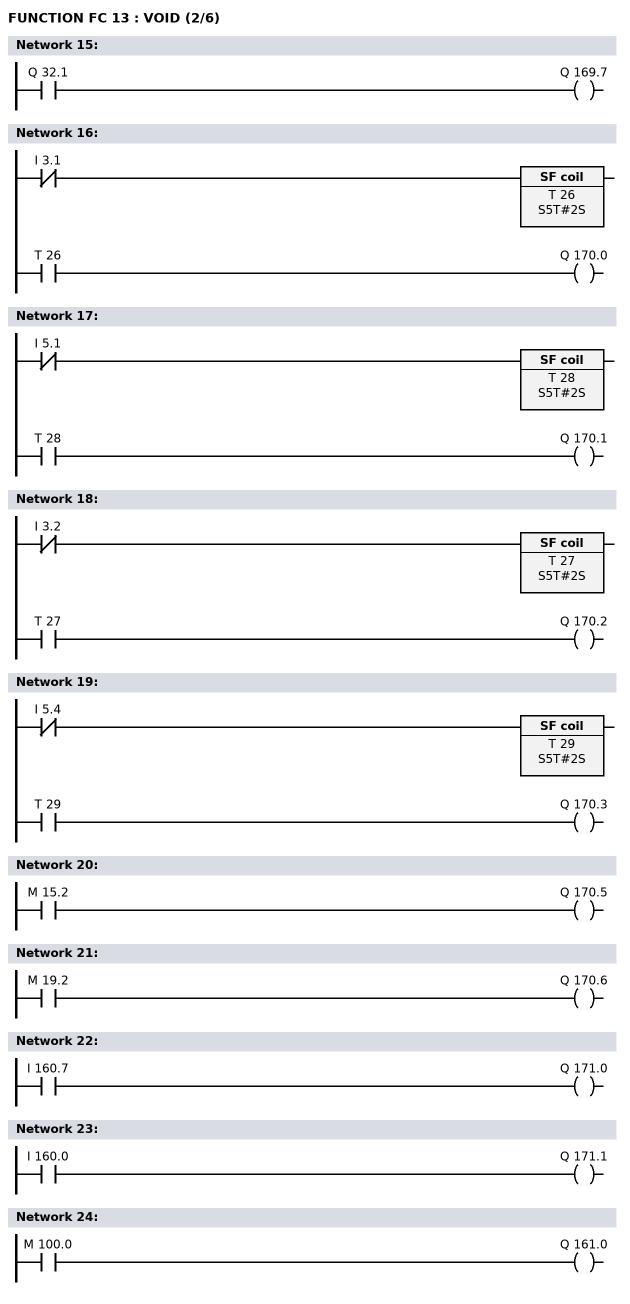

      A     Q     32.1;
      =     Q    169.7;
NETWORK
TITLE =

      AN    I      3.1;
      L     S5T#2S;
      SF    T     26;
      NOP   0;
      NOP   0;
      NOP   0;
      A     T     26;
      =     Q    170.0;
NETWORK
TITLE =

      AN    I      5.1;
      L     S5T#2S;
      SF    T     28;
      NOP   0;
      NOP   0;
      NOP   0;
      A     T     28;
      =     Q    170.1;
NETWORK
TITLE =

      AN    I      3.2;
      L     S5T#2S;
      SF    T     27;
      NOP   0;
      NOP   0;
      NOP   0;
      A     T     27;
      =     Q    170.2;
NETWORK
TITLE =

      AN    I      5.4;
      L     S5T#2S;
      SF    T     29;
      NOP   0;
      NOP   0;
      NOP   0;
      A     T     29;
      =     Q    170.3;
NETWORK
TITLE =

      A     M     15.2;
      =     Q    170.5;
NETWORK
TITLE =

      A     M     19.2;
      =     Q    170.6;
NETWORK
TITLE =

      A     I    160.7;
      =     Q    171.0;
NETWORK
TITLE =

      A     I    160.0;
      =     Q    171.1;
NETWORK
TITLE =

      A     M    100.0;
      =     Q    161.0;
NETWORK
TITLE =
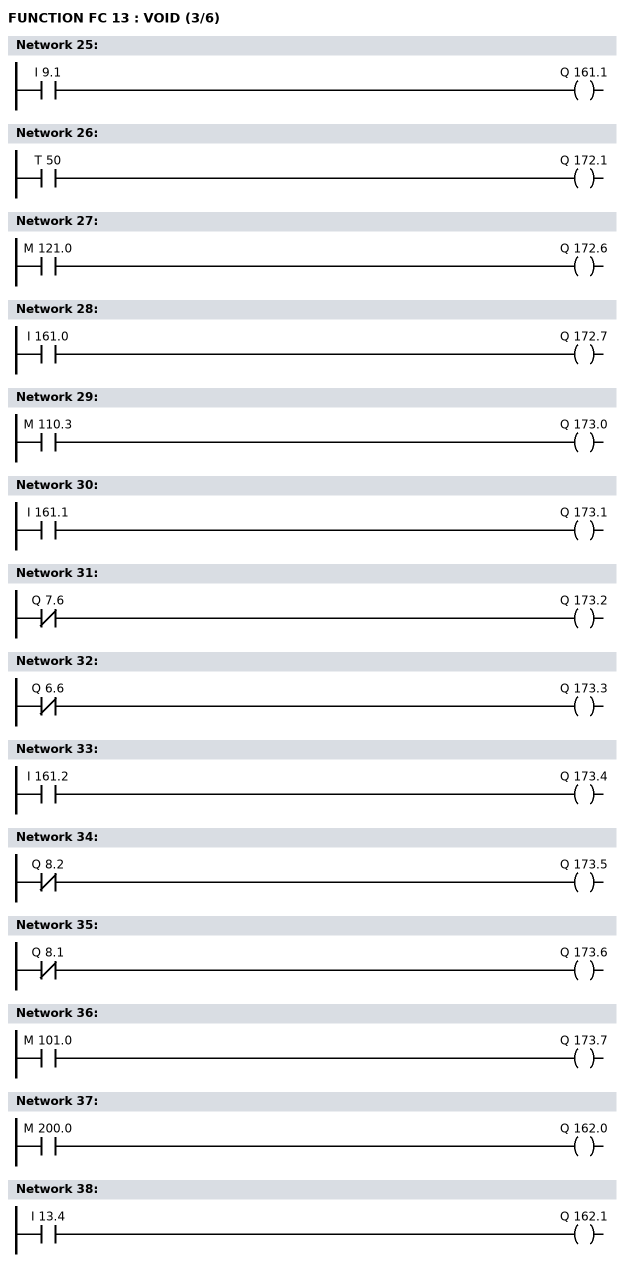

      A     I      9.1;
      =     Q    161.1;
NETWORK
TITLE =

      A     T     50;
      =     Q    172.1;
NETWORK
TITLE =

      A     M    121.0;
      =     Q    172.6;
NETWORK
TITLE =

      A     I    161.0;
      =     Q    172.7;
NETWORK
TITLE =

      A     M    110.3;
      =     Q    173.0;
NETWORK
TITLE =

      A     I    161.1;
      =     Q    173.1;
NETWORK
TITLE =

      AN    Q      7.6;
      =     Q    173.2;
NETWORK
TITLE =

      AN    Q      6.6;
      =     Q    173.3;
NETWORK
TITLE =

      A     I    161.2;
      =     Q    173.4;
NETWORK
TITLE =

      AN    Q      8.2;
      =     Q    173.5;
NETWORK
TITLE =

      AN    Q      8.1;
      =     Q    173.6;
NETWORK
TITLE =

      A     M    101.0;
      =     Q    173.7;
NETWORK
TITLE =

      A     M    200.0;
      =     Q    162.0;
NETWORK
TITLE =

      A     I     13.4;
      =     Q    162.1;
NETWORK
TITLE =
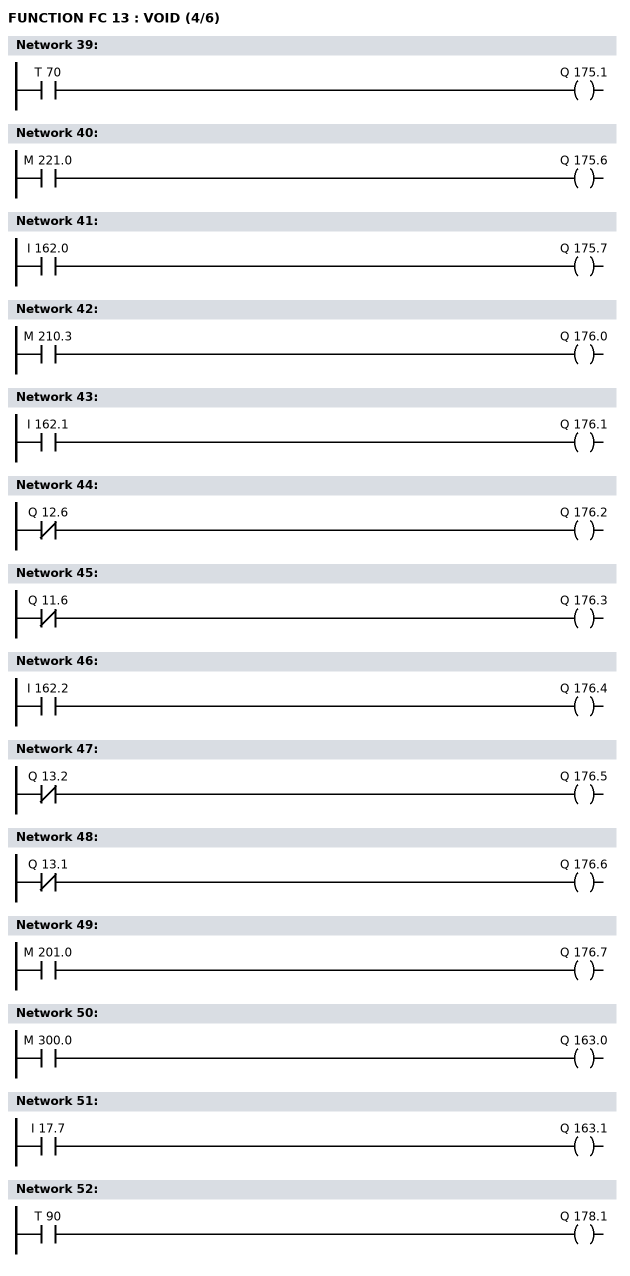

      A     T     70;
      =     Q    175.1;
NETWORK
TITLE =

      A     M    221.0;
      =     Q    175.6;
NETWORK
TITLE =

      A     I    162.0;
      =     Q    175.7;
NETWORK
TITLE =

      A     M    210.3;
      =     Q    176.0;
NETWORK
TITLE =

      A     I    162.1;
      =     Q    176.1;
NETWORK
TITLE =

      AN    Q     12.6;
      =     Q    176.2;
NETWORK
TITLE =

      AN    Q     11.6;
      =     Q    176.3;
NETWORK
TITLE =

      A     I    162.2;
      =     Q    176.4;
NETWORK
TITLE =

      AN    Q     13.2;
      =     Q    176.5;
NETWORK
TITLE =

      AN    Q     13.1;
      =     Q    176.6;
NETWORK
TITLE =

      A     M    201.0;
      =     Q    176.7;
NETWORK
TITLE =

      A     M    300.0;
      =     Q    163.0;
NETWORK
TITLE =

      A     I     17.7;
      =     Q    163.1;
NETWORK
TITLE =

      A     T     90;
      =     Q    178.1;
NETWORK
TITLE =
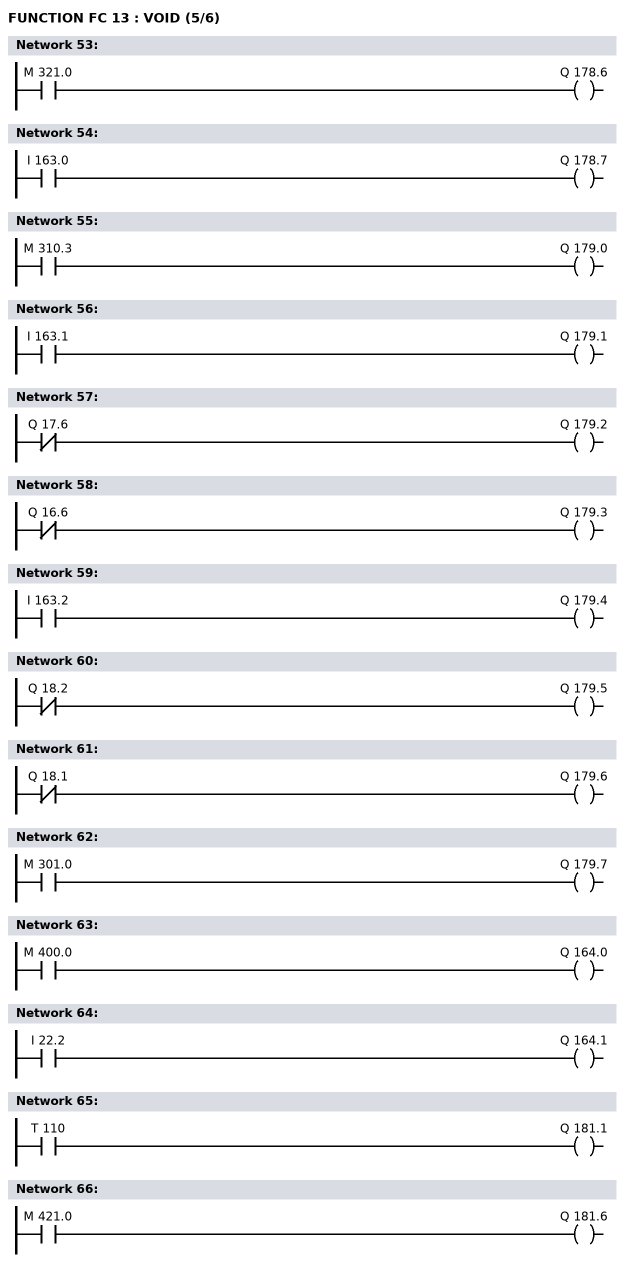

      A     M    321.0;
      =     Q    178.6;
NETWORK
TITLE =

      A     I    163.0;
      =     Q    178.7;
NETWORK
TITLE =

      A     M    310.3;
      =     Q    179.0;
NETWORK
TITLE =

      A     I    163.1;
      =     Q    179.1;
NETWORK
TITLE =

      AN    Q     17.6;
      =     Q    179.2;
NETWORK
TITLE =

      AN    Q     16.6;
      =     Q    179.3;
NETWORK
TITLE =

      A     I    163.2;
      =     Q    179.4;
NETWORK
TITLE =

      AN    Q     18.2;
      =     Q    179.5;
NETWORK
TITLE =

      AN    Q     18.1;
      =     Q    179.6;
NETWORK
TITLE =

      A     M    301.0;
      =     Q    179.7;
NETWORK
TITLE =

      A     M    400.0;
      =     Q    164.0;
NETWORK
TITLE =

      A     I     22.2;
      =     Q    164.1;
NETWORK
TITLE =

      A     T    110;
      =     Q    181.1;
NETWORK
TITLE =

      A     M    421.0;
      =     Q    181.6;
NETWORK
TITLE =
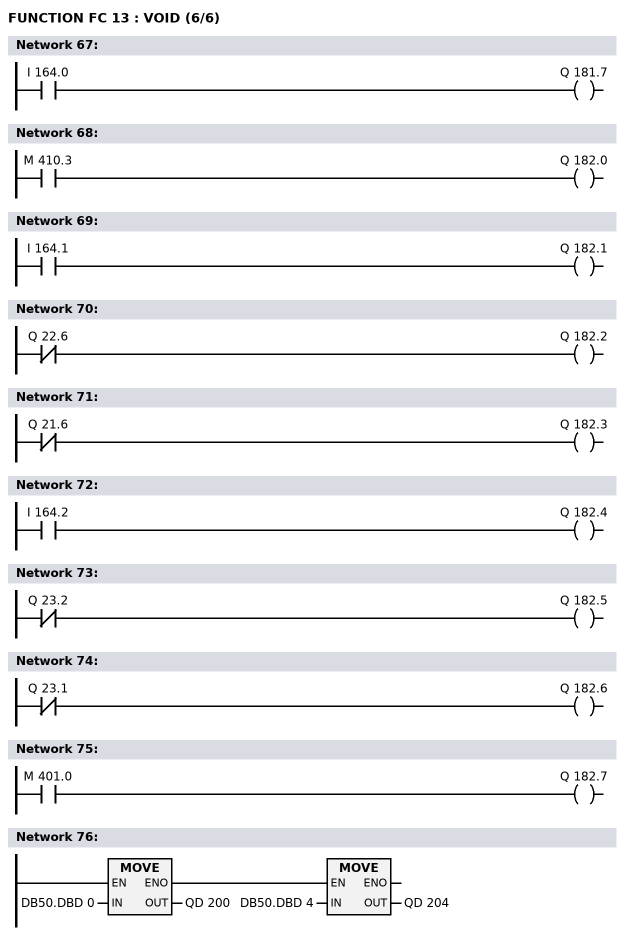

      A     I    164.0;
      =     Q    181.7;
NETWORK
TITLE =

      A     M    410.3;
      =     Q    182.0;
NETWORK
TITLE =

      A     I    164.1;
      =     Q    182.1;
NETWORK
TITLE =

      AN    Q     22.6;
      =     Q    182.2;
NETWORK
TITLE =

      AN    Q     21.6;
      =     Q    182.3;
NETWORK
TITLE =

      A     I    164.2;
      =     Q    182.4;
NETWORK
TITLE =

      AN    Q     23.2;
      =     Q    182.5;
NETWORK
TITLE =

      AN    Q     23.1;
      =     Q    182.6;
NETWORK
TITLE =

      A     M    401.0;
      =     Q    182.7;
NETWORK
TITLE =

      A(    ;
      L     DB50.DBD    0;
      T     QD   200;
      SET   ;
      SAVE  ;
      CLR   ;
      A     BR;
      )     ;
      JNB   M001;
      L     DB50.DBD    4;
      T     QD   204;
M001: NOP   0;
END_FUNCTION

FUNCTION FC 100 : VOID
VERSION : 0.1

BEGIN
NETWORK
TITLE =
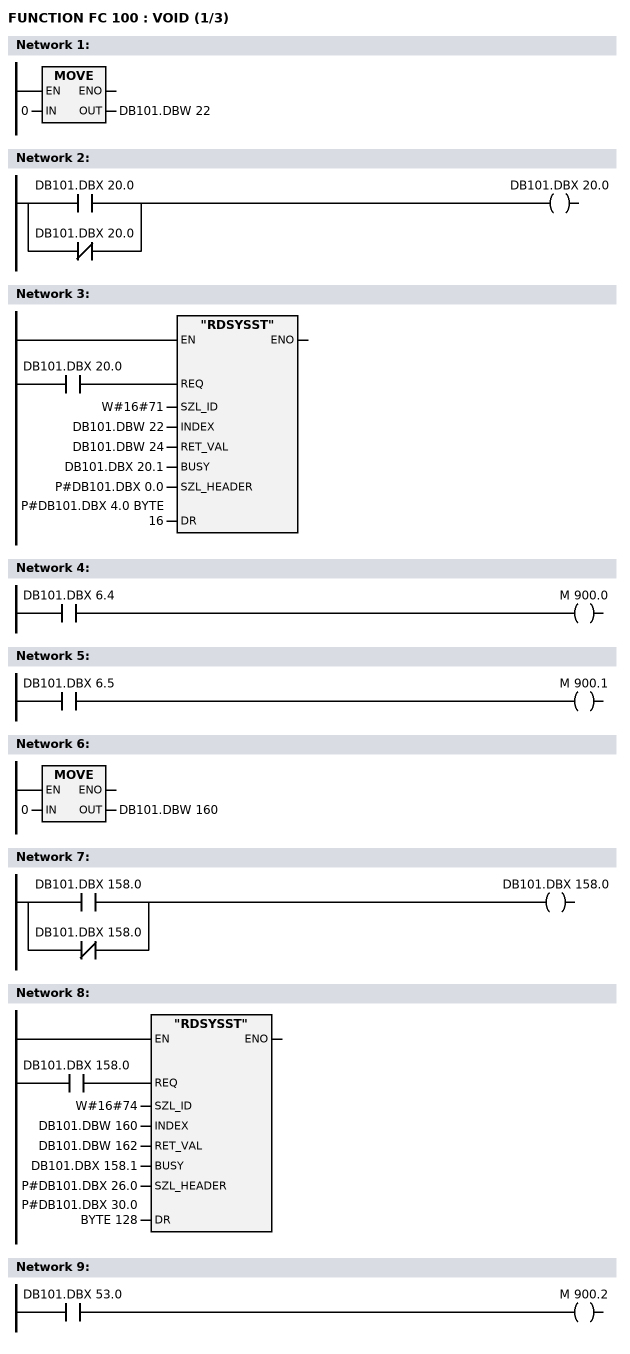

      L     0;
      T     DB101.DBW   22;
      NOP   0;
NETWORK
TITLE =

      O     DB101.DBX   20.0;
      ON    DB101.DBX   20.0;
      =     DB101.DBX   20.0;
NETWORK
TITLE =

      A     DB101.DBX   20.0;
      =     L      0.0;
      BLD   103;
      CALL "RDSYSST" (
           REQ                      := L      0.0,
           SZL_ID                   := W#16#71,
           INDEX                    := DB101.DBW   22,
           RET_VAL                  := DB101.DBW   24,
           BUSY                     := DB101.DBX   20.1,
           SZL_HEADER               := P#DB101.DBX 0.0,
           DR                       := P#DB101.DBX 4.0 BYTE 16);
      NOP   0;
NETWORK
TITLE =

      A     DB101.DBX    6.4;
      =     M    900.0;
NETWORK
TITLE =

      A     DB101.DBX    6.5;
      =     M    900.1;
NETWORK
TITLE =

      L     0;
      T     DB101.DBW  160;
      NOP   0;
NETWORK
TITLE =

      O     DB101.DBX  158.0;
      ON    DB101.DBX  158.0;
      =     DB101.DBX  158.0;
NETWORK
TITLE =

      A     DB101.DBX  158.0;
      =     L      0.0;
      BLD   103;
      CALL "RDSYSST" (
           REQ                      := L      0.0,
           SZL_ID                   := W#16#74,
           INDEX                    := DB101.DBW  160,
           RET_VAL                  := DB101.DBW  162,
           BUSY                     := DB101.DBX  158.1,
           SZL_HEADER               := P#DB101.DBX 26.0,
           DR                       := P#DB101.DBX 30.0 BYTE 128);
      NOP   0;
NETWORK
TITLE =

      A     DB101.DBX   53.0;
      =     M    900.2;
NETWORK
TITLE =
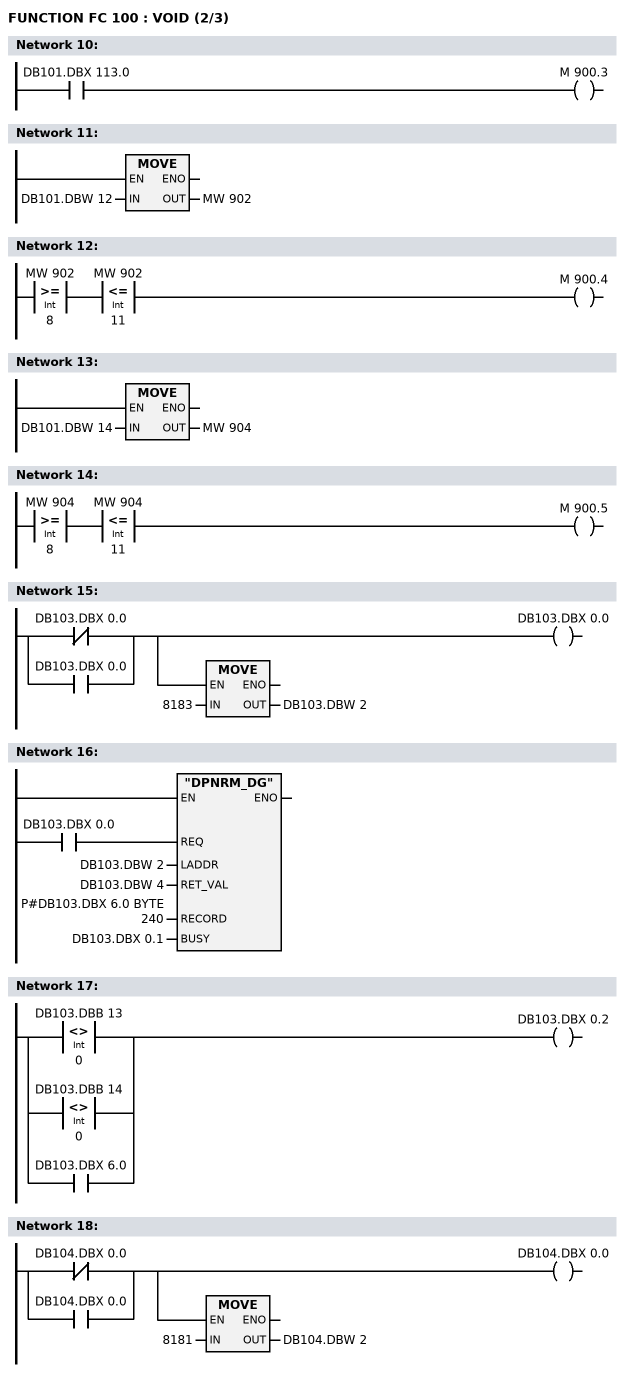

      A     DB101.DBX  113.0;
      =     M    900.3;
NETWORK
TITLE =

      L     DB101.DBW   12;
      T     MW   902;
      NOP   0;
NETWORK
TITLE =

      A(    ;
      L     MW   902;
      L     8;
      >=I   ;
      )     ;
      A(    ;
      L     MW   902;
      L     11;
      <=I   ;
      )     ;
      =     M    900.4;
NETWORK
TITLE =

      L     DB101.DBW   14;
      T     MW   904;
      NOP   0;
NETWORK
TITLE =

      A(    ;
      L     MW   904;
      L     8;
      >=I   ;
      )     ;
      A(    ;
      L     MW   904;
      L     11;
      <=I   ;
      )     ;
      =     M    900.5;
NETWORK
TITLE =

      ON    DB103.DBX    0.0;
      O     DB103.DBX    0.0;
      =     L      0.0;
      A     L      0.0;
      BLD   102;
      =     DB103.DBX    0.0;
      A     L      0.0;
      JNB   M001;
      L     8183;
      T     DB103.DBW    2;
M001: NOP   0;
NETWORK
TITLE =

      A     DB103.DBX    0.0;
      =     L      0.0;
      BLD   103;
      CALL "DPNRM_DG" (
           REQ                      := L      0.0,
           LADDR                    := DB103.DBW    2,
           RET_VAL                  := DB103.DBW    4,
           RECORD                   := P#DB103.DBX 6.0 BYTE 240,
           BUSY                     := DB103.DBX    0.1);
      NOP   0;
NETWORK
TITLE =

      O(    ;
      L     DB103.DBB   13;
      L     0;
      <>I   ;
      )     ;
      O(    ;
      L     DB103.DBB   14;
      L     0;
      <>I   ;
      )     ;
      O     DB103.DBX    6.0;
      =     DB103.DBX    0.2;
NETWORK
TITLE =

      ON    DB104.DBX    0.0;
      O     DB104.DBX    0.0;
      =     L      0.0;
      A     L      0.0;
      BLD   102;
      =     DB104.DBX    0.0;
      A     L      0.0;
      JNB   M002;
      L     8181;
      T     DB104.DBW    2;
M002: NOP   0;
NETWORK
TITLE =
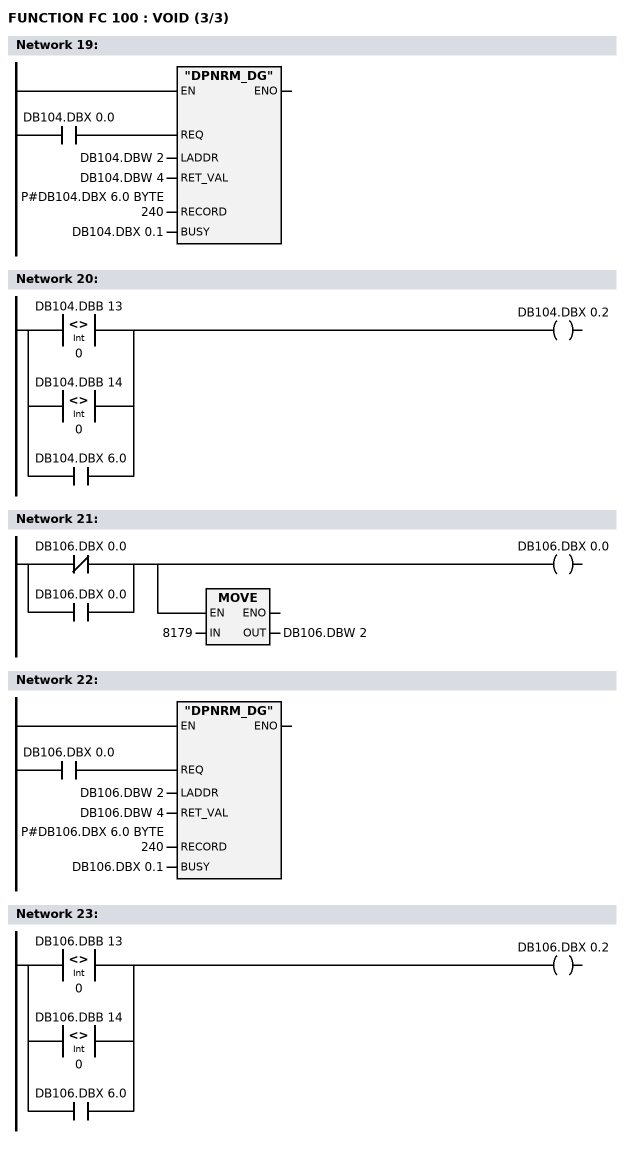

      A     DB104.DBX    0.0;
      =     L      0.0;
      BLD   103;
      CALL "DPNRM_DG" (
           REQ                      := L      0.0,
           LADDR                    := DB104.DBW    2,
           RET_VAL                  := DB104.DBW    4,
           RECORD                   := P#DB104.DBX 6.0 BYTE 240,
           BUSY                     := DB104.DBX    0.1);
      NOP   0;
NETWORK
TITLE =

      O(    ;
      L     DB104.DBB   13;
      L     0;
      <>I   ;
      )     ;
      O(    ;
      L     DB104.DBB   14;
      L     0;
      <>I   ;
      )     ;
      O     DB104.DBX    6.0;
      =     DB104.DBX    0.2;
NETWORK
TITLE =

      ON    DB106.DBX    0.0;
      O     DB106.DBX    0.0;
      =     L      0.0;
      A     L      0.0;
      BLD   102;
      =     DB106.DBX    0.0;
      A     L      0.0;
      JNB   M003;
      L     8179;
      T     DB106.DBW    2;
M003: NOP   0;
NETWORK
TITLE =

      A     DB106.DBX    0.0;
      =     L      0.0;
      BLD   103;
      CALL "DPNRM_DG" (
           REQ                      := L      0.0,
           LADDR                    := DB106.DBW    2,
           RET_VAL                  := DB106.DBW    4,
           RECORD                   := P#DB106.DBX 6.0 BYTE 240,
           BUSY                     := DB106.DBX    0.1);
      NOP   0;
NETWORK
TITLE =

      O(    ;
      L     DB106.DBB   13;
      L     0;
      <>I   ;
      )     ;
      O(    ;
      L     DB106.DBB   14;
      L     0;
      <>I   ;
      )     ;
      O     DB106.DBX    6.0;
      =     DB106.DBX    0.2;
END_FUNCTION

DATA_BLOCK DB 500
VERSION : 0.0

 FB 500
BEGIN
   IN0 := FALSE;
   IN1 := FALSE;
   IN2 := FALSE;
   OUT3 := FALSE;
   OUT4 := FALSE;
   STAT5 := FALSE;
   STAT6 := FALSE;
   STAT7 := FALSE;
   STAT8 := FALSE;
END_DATA_BLOCK

DATA_BLOCK DB 501
VERSION : 0.0

 FB 500
BEGIN
   IN0 := FALSE;
   IN1 := FALSE;
   IN2 := FALSE;
   OUT3 := FALSE;
   OUT4 := FALSE;
   STAT5 := FALSE;
   STAT6 := FALSE;
   STAT7 := FALSE;
   STAT8 := FALSE;
END_DATA_BLOCK

DATA_BLOCK DB 502
VERSION : 0.0

 FB 500
BEGIN
   IN0 := FALSE;
   IN1 := FALSE;
   IN2 := FALSE;
   OUT3 := FALSE;
   OUT4 := FALSE;
   STAT5 := FALSE;
   STAT6 := FALSE;
   STAT7 := FALSE;
   STAT8 := FALSE;
END_DATA_BLOCK

DATA_BLOCK DB 504
VERSION : 0.0

 FB 500
BEGIN
   IN0 := FALSE;
   IN1 := FALSE;
   IN2 := FALSE;
   OUT3 := FALSE;
   OUT4 := FALSE;
   STAT5 := FALSE;
   STAT6 := FALSE;
   STAT7 := FALSE;
   STAT8 := FALSE;
END_DATA_BLOCK

DATA_BLOCK DB 505
VERSION : 0.0

 FB 500
BEGIN
   IN0 := FALSE;
   IN1 := FALSE;
   IN2 := FALSE;
   OUT3 := FALSE;
   OUT4 := FALSE;
   STAT5 := FALSE;
   STAT6 := FALSE;
   STAT7 := FALSE;
   STAT8 := FALSE;
END_DATA_BLOCK

DATA_BLOCK DB 506
VERSION : 0.0

 FB 500
BEGIN
   IN0 := FALSE;
   IN1 := FALSE;
   IN2 := FALSE;
   OUT3 := FALSE;
   OUT4 := FALSE;
   STAT5 := FALSE;
   STAT6 := FALSE;
   STAT7 := FALSE;
   STAT8 := FALSE;
END_DATA_BLOCK

DATA_BLOCK DB 507
VERSION : 0.0

 FB 500
BEGIN
   IN0 := FALSE;
   IN1 := FALSE;
   IN2 := FALSE;
   OUT3 := FALSE;
   OUT4 := FALSE;
   STAT5 := FALSE;
   STAT6 := FALSE;
   STAT7 := FALSE;
   STAT8 := FALSE;
END_DATA_BLOCK

DATA_BLOCK DB 508
VERSION : 0.0

 FB 500
BEGIN
   IN0 := FALSE;
   IN1 := FALSE;
   IN2 := FALSE;
   OUT3 := FALSE;
   OUT4 := FALSE;
   STAT5 := FALSE;
   STAT6 := FALSE;
   STAT7 := FALSE;
   STAT8 := FALSE;
END_DATA_BLOCK

DATA_BLOCK DB 509
VERSION : 0.0

 FB 500
BEGIN
   IN0 := FALSE;
   IN1 := FALSE;
   IN2 := FALSE;
   OUT3 := FALSE;
   OUT4 := FALSE;
   STAT5 := FALSE;
   STAT6 := FALSE;
   STAT7 := FALSE;
   STAT8 := FALSE;
END_DATA_BLOCK

DATA_BLOCK DB 517
VERSION : 0.0

 FB 500
BEGIN
   IN0 := FALSE;
   IN1 := FALSE;
   IN2 := FALSE;
   OUT3 := FALSE;
   OUT4 := FALSE;
   STAT5 := FALSE;
   STAT6 := FALSE;
   STAT7 := FALSE;
   STAT8 := FALSE;
END_DATA_BLOCK

DATA_BLOCK DB 518
VERSION : 0.0

 FB 500
BEGIN
   IN0 := FALSE;
   IN1 := FALSE;
   IN2 := FALSE;
   OUT3 := FALSE;
   OUT4 := FALSE;
   STAT5 := FALSE;
   STAT6 := FALSE;
   STAT7 := FALSE;
   STAT8 := FALSE;
END_DATA_BLOCK

DATA_BLOCK DB 519
VERSION : 0.0

 FB 500
BEGIN
   IN0 := FALSE;
   IN1 := FALSE;
   IN2 := FALSE;
   OUT3 := FALSE;
   OUT4 := FALSE;
   STAT5 := FALSE;
   STAT6 := FALSE;
   STAT7 := FALSE;
   STAT8 := FALSE;
END_DATA_BLOCK

DATA_BLOCK DB 520
VERSION : 0.0

 FB 500
BEGIN
   IN0 := FALSE;
   IN1 := FALSE;
   IN2 := FALSE;
   OUT3 := FALSE;
   OUT4 := FALSE;
   STAT5 := FALSE;
   STAT6 := FALSE;
   STAT7 := FALSE;
   STAT8 := FALSE;
END_DATA_BLOCK

DATA_BLOCK DB 521
VERSION : 0.0

 FB 500
BEGIN
   IN0 := FALSE;
   IN1 := FALSE;
   IN2 := FALSE;
   OUT3 := FALSE;
   OUT4 := FALSE;
   STAT5 := FALSE;
   STAT6 := FALSE;
   STAT7 := FALSE;
   STAT8 := FALSE;
END_DATA_BLOCK

DATA_BLOCK DB 522
VERSION : 0.0

 FB 500
BEGIN
   IN0 := FALSE;
   IN1 := FALSE;
   IN2 := FALSE;
   OUT3 := FALSE;
   OUT4 := FALSE;
   STAT5 := FALSE;
   STAT6 := FALSE;
   STAT7 := FALSE;
   STAT8 := FALSE;
END_DATA_BLOCK

DATA_BLOCK DB 523
VERSION : 0.0

 FB 500
BEGIN
   IN0 := FALSE;
   IN1 := FALSE;
   IN2 := FALSE;
   OUT3 := FALSE;
   OUT4 := FALSE;
   STAT5 := FALSE;
   STAT6 := FALSE;
   STAT7 := FALSE;
   STAT8 := FALSE;
END_DATA_BLOCK

DATA_BLOCK DB 524
VERSION : 0.0

 FB 500
BEGIN
   IN0 := FALSE;
   IN1 := FALSE;
   IN2 := FALSE;
   OUT3 := FALSE;
   OUT4 := FALSE;
   STAT5 := FALSE;
   STAT6 := FALSE;
   STAT7 := FALSE;
   STAT8 := FALSE;
END_DATA_BLOCK

ORGANIZATION_BLOCK OB 1
VERSION : 0.1


VAR_TEMP
  TEMP0 : BYTE ;
  TEMP1 : BYTE ;
  TEMP2 : BYTE ;
  TEMP3 : BYTE ;
  TEMP4 : BYTE ;
  TEMP5 : BYTE ;
  TEMP6 : INT ;
  TEMP7 : INT ;
  TEMP8 : INT ;
  TEMP9 : DATE_AND_TIME ;
END_VAR
BEGIN
NETWORK
TITLE =
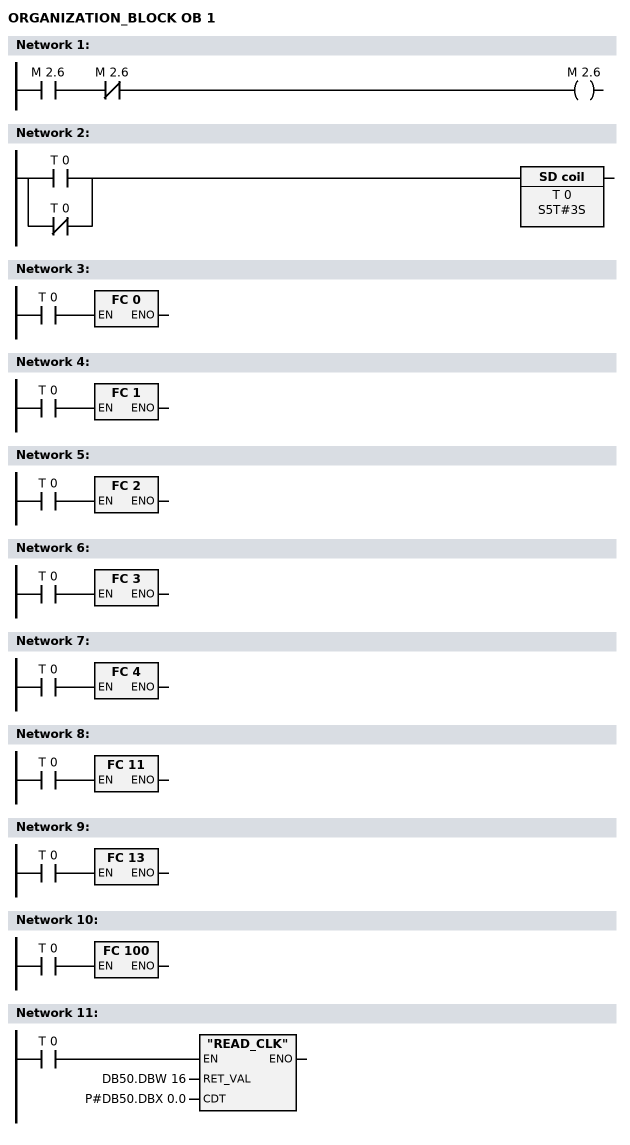

      A     M      2.6;
      AN    M      2.6;
      =     M      2.6;
NETWORK
TITLE =

      A(    ;
      O     T      0;
      ON    T      0;
      )     ;
      L     S5T#3S;
      SD    T      0;
      NOP   0;
      NOP   0;
      NOP   0;
      NOP   0;
NETWORK
TITLE =

      A     T      0;
      JNB   M001;
      CALL FC     0 ;
M001: NOP   0;
NETWORK
TITLE =

      A     T      0;
      JNB   M002;
      CALL FC     1 ;
M002: NOP   0;
NETWORK
TITLE =

      A     T      0;
      JNB   M003;
      CALL FC     2 ;
M003: NOP   0;
NETWORK
TITLE =

      A     T      0;
      JNB   M004;
      CALL FC     3 ;
M004: NOP   0;
NETWORK
TITLE =

      A     T      0;
      JNB   M005;
      CALL FC     4 ;
M005: NOP   0;
NETWORK
TITLE =

      A     T      0;
      JNB   M006;
      CALL FC    11 ;
M006: NOP   0;
NETWORK
TITLE =

      A     T      0;
      JNB   M007;
      CALL FC    13 ;
M007: NOP   0;
NETWORK
TITLE =

      A     T      0;
      JNB   M008;
      CALL FC   100 ;
M008: NOP   0;
NETWORK
TITLE =

      A     T      0;
      JNB   M009;
      CALL "READ_CLK" (
           RET_VAL                  := DB50.DBW   16,
           CDT                      := P#DB50.DBX 0.0);
M009: NOP   0;
END_ORGANIZATION_BLOCK

ORGANIZATION_BLOCK OB 35
VERSION : 0.1


VAR_TEMP
  TEMP0 : BYTE ;
  TEMP1 : BYTE ;
  TEMP2 : BYTE ;
  TEMP3 : BYTE ;
  TEMP4 : BYTE ;
  TEMP5 : BYTE ;
  TEMP6 : WORD ;
  TEMP7 : INT ;
  TEMP8 : INT ;
  TEMP9 : DATE_AND_TIME ;
END_VAR
BEGIN
END_ORGANIZATION_BLOCK

ORGANIZATION_BLOCK OB 70
VERSION : 0.1


VAR_TEMP
  TEMP0 : BYTE ;
  TEMP1 : BYTE ;
  TEMP2 : BYTE ;
  TEMP3 : BYTE ;
  TEMP4 : WORD ;
  TEMP5 : WORD ;
  TEMP6 : WORD ;
  TEMP7 : WORD ;
  TEMP8 : DATE_AND_TIME ;
END_VAR
BEGIN
NETWORK
TITLE =

      AN    M      3.7;
      =     M      3.7;
END_ORGANIZATION_BLOCK

ORGANIZATION_BLOCK OB 72
VERSION : 0.1


VAR_TEMP
  TEMP0 : BYTE ;
  TEMP1 : BYTE ;
  TEMP2 : BYTE ;
  TEMP3 : BYTE ;
  TEMP4 : WORD ;
  TEMP5 : WORD ;
  TEMP6 : WORD ;
  TEMP7 : WORD ;
  TEMP8 : DATE_AND_TIME ;
END_VAR
BEGIN
NETWORK
TITLE =

      A     M      3.7;
      =     M      3.7;
END_ORGANIZATION_BLOCK

ORGANIZATION_BLOCK OB 81
VERSION : 0.1


VAR_TEMP
  TEMP0 : BYTE ;
  TEMP1 : BYTE ;
  TEMP2 : BYTE ;
  TEMP3 : BYTE ;
  TEMP4 : BYTE ;
  TEMP5 : BYTE ;
  TEMP6 : WORD ;
  TEMP7 : BYTE ;
  TEMP8 : BYTE ;
  TEMP9 : BYTE ;
  TEMP10 : BYTE ;
  TEMP11 : DATE_AND_TIME ;
END_VAR
BEGIN
NETWORK
TITLE =

      AN    M      3.7;
      =     M      3.7;
END_ORGANIZATION_BLOCK

ORGANIZATION_BLOCK OB 82
VERSION : 0.1


VAR_TEMP
  TEMP0 : BYTE ;
  TEMP1 : BYTE ;
  TEMP2 : BYTE ;
  TEMP3 : BYTE ;
  TEMP4 : BYTE ;
  TEMP5 : BYTE ;
  TEMP6 : WORD ;
  TEMP7 : BOOL ;
  TEMP8 : BOOL ;
  TEMP9 : BOOL ;
  TEMP10 : BOOL ;
  TEMP11 : BOOL ;
  TEMP12 : BOOL ;
  TEMP13 : BOOL ;
  TEMP14 : BOOL ;
  TEMP15 : BYTE ;
  TEMP16 : BOOL ;
  TEMP17 : BOOL ;
  TEMP18 : BOOL ;
  TEMP19 : BOOL ;
  TEMP20 : BOOL ;
  TEMP21 : BOOL ;
  TEMP22 : BOOL ;
  TEMP23 : BOOL ;
  TEMP24 : BOOL ;
  TEMP25 : BOOL ;
  TEMP26 : BOOL ;
  TEMP27 : BOOL ;
  TEMP28 : BOOL ;
  TEMP29 : BOOL ;
  TEMP30 : BOOL ;
  TEMP31 : BOOL ;
  TEMP32 : DATE_AND_TIME ;
END_VAR
BEGIN
NETWORK
TITLE =

      AN    M      3.7;
      =     M      3.7;
END_ORGANIZATION_BLOCK

ORGANIZATION_BLOCK OB 83
VERSION : 0.1


VAR_TEMP
  TEMP0 : BYTE ;
  TEMP1 : BYTE ;
  TEMP2 : BYTE ;
  TEMP3 : BYTE ;
  TEMP4 : BYTE ;
  TEMP5 : BYTE ;
  TEMP6 : WORD ;
  TEMP7 : INT ;
  TEMP8 : WORD ;
  TEMP9 : DATE_AND_TIME ;
END_VAR
BEGIN
NETWORK
TITLE =

      AN    M      3.7;
      =     M      3.7;
END_ORGANIZATION_BLOCK

ORGANIZATION_BLOCK OB 85
VERSION : 0.1


VAR_TEMP
  TEMP0 : BYTE ;
  TEMP1 : BYTE ;
  TEMP2 : BYTE ;
  TEMP3 : BYTE ;
  TEMP4 : BYTE ;
  TEMP5 : BYTE ;
  TEMP6 : INT ;
  TEMP7 : BYTE ;
  TEMP8 : BYTE ;
  TEMP9 : BYTE ;
  TEMP10 : BYTE ;
  TEMP11 : DATE_AND_TIME ;
END_VAR
BEGIN
NETWORK
TITLE =

      AN    M      3.7;
      =     M      3.7;
END_ORGANIZATION_BLOCK

ORGANIZATION_BLOCK OB 86
VERSION : 0.1


VAR_TEMP
  TEMP0 : BYTE ;
  TEMP1 : BYTE ;
  TEMP2 : BYTE ;
  TEMP3 : BYTE ;
  TEMP4 : BYTE ;
  TEMP5 : BYTE ;
  TEMP6 : WORD ;
  TEMP7 : ARRAY  [0 .. 31 ] OF BOOL ;
  TEMP8 : DATE_AND_TIME ;
END_VAR
BEGIN
NETWORK
TITLE =

      AN    M      3.7;
      =     M      3.7;
END_ORGANIZATION_BLOCK

ORGANIZATION_BLOCK OB 87
VERSION : 0.1


VAR_TEMP
  TEMP0 : BYTE ;
  TEMP1 : BYTE ;
  TEMP2 : BYTE ;
  TEMP3 : BYTE ;
  TEMP4 : BYTE ;
  TEMP5 : BYTE ;
  TEMP6 : WORD ;
  TEMP7 : DWORD ;
  TEMP8 : DATE_AND_TIME ;
END_VAR
BEGIN
NETWORK
TITLE =

      AN    M      3.7;
      =     M      3.7;
END_ORGANIZATION_BLOCK

ORGANIZATION_BLOCK OB 100
VERSION : 0.1


VAR_TEMP
  TEMP0 : BYTE ;
  TEMP1 : BYTE ;
  TEMP2 : BYTE ;
  TEMP3 : BYTE ;
  TEMP4 : BYTE ;
  TEMP5 : BYTE ;
  TEMP6 : WORD ;
  TEMP7 : DWORD ;
  TEMP8 : DATE_AND_TIME ;
END_VAR
BEGIN
END_ORGANIZATION_BLOCK

ORGANIZATION_BLOCK OB 122
VERSION : 0.1


VAR_TEMP
  TEMP0 : BYTE ;
  TEMP1 : BYTE ;
  TEMP2 : BYTE ;
  TEMP3 : BYTE ;
  TEMP4 : BYTE ;
  TEMP5 : BYTE ;
  TEMP6 : WORD ;
  TEMP7 : WORD ;
  TEMP8 : WORD ;
  TEMP9 : DATE_AND_TIME ;
END_VAR
BEGIN
NETWORK
TITLE =

      AN    M      3.7;
      =     M      3.7;
END_ORGANIZATION_BLOCK
